Staubli VAL3: initCombo.pgx

public program initCombo(utCombo& x_utCombo[], string x_sPage, string x_sId)
begin
  x_utCombo.Common.sPage=x_sPage
  x_utCombo.Common.sID=x_sId
  userPageBind(x_utCombo.Common.sPage,x_utCombo.Common.sID,"options",x_utCombo.Common.sItem,size(x_utCombo.Common.sItem),"r")
  userPageBind(x_utCombo.Common.sPage,x_utCombo.Common.sID,"value",x_utCombo.Common.sValue,1,"rw")
end
